(* IEC 61131-3 sources: PLC_ST_Simulator/, 2 files *)

(* ---- Saege_CODESYS.st ---- *)
VAR_GLOBAL
    E0  : BOOL;  (* S0  Rohr an Anschlag 1 *)
    E1  : BOOL;  (* S1  Rohr an Anschlag 2 *)
    E2  : BOOL;  (* S2  gespannt *)
    E3  : BOOL;  (* S3  entspannt *)
    E4  : BOOL;  (* S4  Säge oben *)
    E5  : BOOL;  (* S5  Säge unten *)
    E6  : BOOL;  (* S6  Anschlag 1 oben *)
    E7  : BOOL;  (* S7  Anschlag 1 unten *)
    E8  : BOOL;  (* S8  EIN *)
    E9  : BOOL;  (* S9  AUS, Öffner *)
    E10 : BOOL;  (* S10 Start *)
    E11 : BOOL;  (* S11 Stopp, Öffner *)
    E12 : BOOL;  (* S12 Anschlag 2 oben *)
    E13 : BOOL;  (* S13 Anschlag 2 unten *)
    E14 : BOOL;  (* S14 dickes Rohr *)
    E15 : BOOL;  (* S15 dünnes Rohr *)
    WST_ABTRANSPORT      : BOOL;  (* B1 *)
    mot_schutz_saege     : BOOL;  (* F1..F5 Öffner *)
    mot_schutz_rolle1    : BOOL;
    mot_schutz_rolle2    : BOOL;
    mot_schutz_anschlag1 : BOOL;
    mot_schutz_anschlag2 : BOOL;

    SAEGE_RUNTER     : BOOL;  (* A1 *)
    SAEGE_HOCH       : BOOL;  (* A2 *)
    SPANNEN          : BOOL;  (* A3 *)
    ENTSPANNEN       : BOOL;  (* A4 *)
    SAEGE_ANTRIEB    : BOOL;  (* K1 *)
    ROLLE_1          : BOOL;  (* K2 *)
    ROLLE_2          : BOOL;  (* K3 *)
    ANSCHLAG1_HOCH   : BOOL;  (* K4 *)
    ANSCHLAG1_RUNTER : BOOL;  (* K5 *)
    ANSCHLAG2_HOCH   : BOOL;  (* K6 *)
    ANSCHLAG2_RUNTER : BOOL;  (* K7 *)
END_VAR

FUNCTION_BLOCK FB_Betriebsart
VAR_OUTPUT
    xEin      : BOOL;
    xAuto     : BOOL;
    xStoerung : BOOL;
END_VAR

xStoerung := NOT (mot_schutz_saege AND mot_schutz_rolle1 AND mot_schutz_rolle2
                  AND mot_schutz_anschlag1 AND mot_schutz_anschlag2);

IF E8 THEN xEin := TRUE;END_IF
IF NOT E9 OR xStoerung THEN xEin := FALSE; END_IF

(* Stopp: laufendes Rohr wird fertig bearbeitet *)
IF E10 AND xEin THEN xAuto := TRUE; END_IF
IF NOT E11 OR NOT xEin THEN xAuto := FALSE; END_IF
END_FUNCTION_BLOCK

PROGRAM SFC_Saege
VAR_INPUT
    xAuto      : BOOL;
    xB1_Flanke : BOOL;
    xReset     : BOOL;   (* zurueck in Grundstellung S1 *)
END_VAR
VAR
    iStep     : INT := 1;
    iStepOld  : INT := 0;
    xNeu      : BOOL;    (* Schritt wurde in diesem Zyklus betreten *)
    xDuenn    : BOOL;
    xDick     : BOOL;
    iSoll     : INT;
    iZaehler  : INT;
    xK1, xK2, xK3, xK5, xK7 : BOOL;
    xAbtransport : BOOL;
    xA1, xA2, xA3, xA4 : BOOL;
END_VAR

(* Reset *)
IF xReset THEN
    iStep    := 1;
    iZaehler := 0;
    xDuenn   := FALSE;
    xDick    := FALSE;
END_IF

xNeu     := (iStep <> iStepOld);
iStepOld := iStep;
(* Start *)
IF xNeu THEN
    CASE iStep OF
        2:  (* ACT_Rohrtyp *)
            xDuenn := E15;
            xDick  := E14 AND NOT E15;
            IF xDuenn THEN iSoll := 4; ELSE iSoll := 3; END_IF
        10: (* ACT_Zaehlen *)
            iZaehler := iZaehler + 1;
        11: (* ACT_Ruecksetzen *)
            iZaehler := 0;
            xDuenn   := FALSE;
            xDick    := FALSE;
    END_CASE
END_IF

(*Schrittekette *)
CASE iStep OF
    1:  IF xAuto AND E3 AND E4 AND E6 AND E12 AND (E14 OR E15) THEN iStep := 2;  END_IF
    2:  IF xDuenn THEN iStep := 3;
        ELSIF xDick THEN iStep := 4; END_IF
    3:  IF E7  THEN iStep := 5; END_IF
    4:  IF E13 THEN iStep := 5; END_IF
    5:  IF (xDuenn AND E0) OR (xDick AND E1) THEN iStep := 6; END_IF
    6:  IF E2  THEN iStep := 7; END_IF
    7:  IF E5  THEN iStep := 8; END_IF
    8:  IF E4  THEN iStep := 9; END_IF
    9:  IF E3  THEN iStep := 10; END_IF
    10: IF WST_ABTRANSPORT AND E6 AND E12 THEN
            IF iZaehler < iSoll THEN
                IF xDuenn THEN iStep := 3; ELSE iStep := 4; END_IF
            ELSE
                iStep := 11;
            END_IF
        END_IF
    11: IF xB1_Flanke THEN iStep := 1; END_IF
END_CASE

(* Schrittverriegelungen*)
xK1          := (iStep = 7) OR (iStep = 8);
xK2          := (iStep = 5) OR (iStep = 11);
xK3          := (iStep = 5) OR (iStep = 10) OR (iStep = 11);
xK5          := (iStep = 3);
xK7          := (iStep = 4);
xA1          := (iStep = 7);
xA2          := (iStep = 8);
xA3          := (iStep = 6);
xA4          := (iStep = 9);
xAbtransport := (iStep = 10);
END_PROGRAM

PROGRAM PRG_Ausgaenge
VAR_INPUT
    xFreigabe : BOOL;
END_VAR

ROLLE_1          := xFreigabe AND SFC_Saege.xK2 AND E3;
ROLLE_2          := xFreigabe AND SFC_Saege.xK3;
SPANNEN          := xFreigabe AND SFC_Saege.xA3 AND NOT SFC_Saege.xA4;
ENTSPANNEN       := xFreigabe AND SFC_Saege.xA4 AND E4;
SAEGE_ANTRIEB    := xFreigabe AND SFC_Saege.xK1 AND E2;
SAEGE_RUNTER     := xFreigabe AND SFC_Saege.xA1 AND E2 AND NOT SFC_Saege.xA2;
SAEGE_HOCH       := xFreigabe AND SFC_Saege.xA2;
ANSCHLAG1_HOCH   := xFreigabe AND SFC_Saege.xAbtransport AND SFC_Saege.xDuenn;
ANSCHLAG2_HOCH   := xFreigabe AND SFC_Saege.xAbtransport AND SFC_Saege.xDick;
ANSCHLAG1_RUNTER := xFreigabe AND SFC_Saege.xK5 AND NOT ANSCHLAG1_HOCH;
ANSCHLAG2_RUNTER := xFreigabe AND SFC_Saege.xK7 AND NOT ANSCHLAG2_HOCH;
END_PROGRAM

PROGRAM PLC_PRG
VAR
    fbBetriebsart : FB_Betriebsart;
    rtB1          : R_TRIG;
END_VAR

fbBetriebsart();
rtB1(CLK := WST_ABTRANSPORT);

SFC_Saege(xAuto := fbBetriebsart.xAuto, xB1_Flanke := rtB1.Q, xReset := NOT fbBetriebsart.xEin);

PRG_Ausgaenge(xFreigabe := fbBetriebsart.xEin AND NOT fbBetriebsart.xStoerung);
END_PROGRAM

(* ---- Saege_Anlage.st ---- *)
(* ============================================================
   Anlagenmodell Rohrsäge  –  läuft im Simulator in jedem Zyklus
   VOR dem SPS-Programm und bildet die Sensoren (E0..E15, B1)
   aus den Ausgängen (A1..A4, K1..K7) nach.

   Geometrie (mm, ab Sägeblatt):  Anschlag 1 = 300, Anschlag 2 = 500,
   Lichtschranke B1 = 1500.  Rohrlänge 1700 mm.
   ============================================================ *)

PROGRAM SIM_Saege
VAR_INPUT
    xNaechstesDick : BOOL := FALSE;   (* Typ des nächsten Rohres *)
    xNachladen     : BOOL := TRUE;    (* automatisch neues Rohr auflegen *)
END_VAR
VAR_OUTPUT
    iSchnitte      : INT;             (* Anzahl Schnitte gesamt *)
    iAbtransport   : INT;             (* Teile, die die Anlage verlassen haben *)
    iRohre         : INT;             (* aufgelegte Rohre *)
    xKollision     : BOOL;            (* mechanische Kollision erkannt *)
    sKollision     : STRING;
END_VAR
VAR CONSTANT
    POS_A1   : REAL := 300.0;
    POS_A2   : REAL := 500.0;
    POS_B1   : REAL := 1500.0;
    ROHR_LEN : REAL := 1700.0;
    V_ROLLE  : REAL := 0.5;     (* mm/ms *)
    V_SAEGE  : REAL := 0.1;     (* %/ms  -> 1 s Hub *)
    V_SPANN  : REAL := 0.4;     (* %/ms  -> 250 ms *)
    V_ANSCHL : REAL := 0.25;    (* %/ms  -> 400 ms *)
    MAX_TEILE : INT := 8;
END_VAR
VAR
    xInit      : BOOL;
    tLast      : TIME;
    dt         : REAL;
    rSaege     : REAL := 100.0;  (* 100 = oben, 0 = unten *)
    rSpann     : REAL := 0.0;    (* 0 = entspannt, 100 = gespannt *)
    rAnschlag1 : REAL := 0.0;    (* 0 = oben, 100 = unten *)
    rAnschlag2 : REAL := 0.0;
    xRohrDick  : BOOL;
    rRohrFront : REAL;           (* Rohranfang hinter dem Sägeblatt *)
    rRohrLen   : REAL;           (* Restlänge auf der Zuführung *)
    aFront     : ARRAY[1..8] OF REAL;   (* abgesägte Teile auf Rollenbahn 2 *)
    aLen       : ARRAY[1..8] OF REAL;
    nTeile     : INT;
    xGeschnitten : BOOL;
    tonLaden   : TON;
    i, k       : INT;
    rWeg, rHinten : REAL;
END_VAR

(* ---------- Initialisierung beim ersten Zyklus ---------- *)
IF NOT xInit THEN
    xInit := TRUE;
    tLast := TIME();
    E9 := TRUE;  E11 := TRUE;   (* Öffner nicht betätigt *)
    mot_schutz_saege := TRUE;  mot_schutz_rolle1 := TRUE;  mot_schutz_rolle2 := TRUE;
    mot_schutz_anschlag1 := TRUE;  mot_schutz_anschlag2 := TRUE;
END_IF
dt := TIME_TO_REAL(TIME() - tLast);
tLast := TIME();

(* ---------- Säge ---------- *)
IF SAEGE_RUNTER AND NOT SAEGE_HOCH THEN
    rSaege := MAX(0.0, rSaege - V_SAEGE * dt);
ELSIF SAEGE_HOCH AND NOT SAEGE_RUNTER THEN
    rSaege := MIN(100.0, rSaege + V_SAEGE * dt);
END_IF
IF rSaege < 60.0 AND rRohrLen > 0.0 AND NOT SAEGE_ANTRIEB AND NOT xKollision THEN
    xKollision := TRUE;  sKollision := 'Säge fährt ohne Antrieb ins Rohr';
END_IF
IF rSaege < 60.0 AND rRohrLen > 0.0 AND rSpann < 100.0 AND NOT xKollision THEN
    xKollision := TRUE;  sKollision := 'Sägen ohne gespanntes Rohr';
END_IF

(* ---------- Spannbacken ---------- *)
IF SPANNEN AND NOT ENTSPANNEN THEN
    rSpann := MIN(100.0, rSpann + V_SPANN * dt);
ELSIF ENTSPANNEN AND NOT SPANNEN THEN
    rSpann := MAX(0.0, rSpann - V_SPANN * dt);
END_IF

(* ---------- Längenanschläge ---------- *)
IF ANSCHLAG1_RUNTER AND NOT ANSCHLAG1_HOCH THEN rAnschlag1 := MIN(100.0, rAnschlag1 + V_ANSCHL * dt);
ELSIF ANSCHLAG1_HOCH AND NOT ANSCHLAG1_RUNTER THEN rAnschlag1 := MAX(0.0, rAnschlag1 - V_ANSCHL * dt); END_IF
IF ANSCHLAG2_RUNTER AND NOT ANSCHLAG2_HOCH THEN rAnschlag2 := MIN(100.0, rAnschlag2 + V_ANSCHL * dt);
ELSIF ANSCHLAG2_HOCH AND NOT ANSCHLAG2_RUNTER THEN rAnschlag2 := MAX(0.0, rAnschlag2 - V_ANSCHL * dt); END_IF

(* Anschlag fährt auf ein Teil, das unter ihm liegt? *)
FOR i := 1 TO nTeile DO
    rHinten := aFront[i] - aLen[i];
    IF ANSCHLAG1_RUNTER AND rHinten < POS_A1 - 1.0 AND aFront[i] > POS_A1 + 1.0 AND NOT xKollision THEN
        xKollision := TRUE;  sKollision := 'Anschlag 1 fährt auf ein Teil';
    END_IF
    IF ANSCHLAG2_RUNTER AND rHinten < POS_A2 - 1.0 AND aFront[i] > POS_A2 + 1.0 AND NOT xKollision THEN
        xKollision := TRUE;  sKollision := 'Anschlag 2 fährt auf ein Teil';
    END_IF
END_FOR

IF ANSCHLAG1_RUNTER AND rRohrLen > 0.0 AND rRohrFront > POS_A1 + 1.0 AND NOT xKollision THEN
    xKollision := TRUE;  sKollision := 'Anschlag 1 fährt auf das Rohr';
END_IF
IF ANSCHLAG2_RUNTER AND rRohrLen > 0.0 AND rRohrFront > POS_A2 + 1.0 AND NOT xKollision THEN
    xKollision := TRUE;  sKollision := 'Anschlag 2 fährt auf das Rohr';
END_IF

(* ---------- Rohr auf der Zuführung (Rollenbahn 1) ---------- *)
IF ROLLE_1 AND rRohrLen > 0.0 THEN
    IF rSpann > 0.0 THEN
        IF NOT xKollision THEN xKollision := TRUE; sKollision := 'Vorschub gegen gespanntes Rohr'; END_IF
    ELSE
        rWeg := V_ROLLE * dt;
        rRohrFront := rRohrFront + rWeg;
        IF rAnschlag1 > 0.0 AND rRohrFront - rWeg <= POS_A1 + 0.01 THEN rRohrFront := MIN(rRohrFront, POS_A1); END_IF
        IF rAnschlag2 > 0.0 AND rRohrFront - rWeg <= POS_A2 + 0.01 THEN rRohrFront := MIN(rRohrFront, POS_A2); END_IF
        (* Rohrende hat die Säge passiert -> Reststück auf Rollenbahn 2 *)
        IF rRohrFront >= rRohrLen AND nTeile < MAX_TEILE THEN
            nTeile := nTeile + 1;
            aFront[nTeile] := rRohrFront;  aLen[nTeile] := rRohrLen;
            rRohrLen := 0.0;  rRohrFront := 0.0;
        END_IF
    END_IF
END_IF

(* ---------- Schnitt ---------- *)
IF SAEGE_ANTRIEB AND rSaege <= 0.0 AND rSpann >= 100.0 AND NOT xGeschnitten AND rRohrFront > 0.0 AND nTeile < MAX_TEILE THEN
    xGeschnitten := TRUE;
    iSchnitte := iSchnitte + 1;
    nTeile := nTeile + 1;
    aFront[nTeile] := rRohrFront;  aLen[nTeile] := rRohrFront;
    rRohrLen := rRohrLen - rRohrFront;
    rRohrFront := 0.0;
END_IF
IF rSaege >= 100.0 THEN xGeschnitten := FALSE; END_IF

(* ---------- Teile auf Rollenbahn 2 ---------- *)
IF ROLLE_2 THEN
    rWeg := V_ROLLE * dt;
    FOR i := 1 TO nTeile DO
        aFront[i] := aFront[i] + rWeg;
        IF rAnschlag1 > 0.0 AND aFront[i] - rWeg <= POS_A1 + 0.01 THEN aFront[i] := MIN(aFront[i], POS_A1); END_IF
        IF rAnschlag2 > 0.0 AND aFront[i] - rWeg <= POS_A2 + 0.01 THEN aFront[i] := MIN(aFront[i], POS_A2); END_IF
    END_FOR
END_IF
(* Teile, die die Rollenbahn verlassen haben, entfernen *)
i := 1;
WHILE i <= nTeile DO
    IF aFront[i] - aLen[i] > POS_B1 + 300.0 THEN
        FOR k := i TO nTeile - 1 DO
            aFront[k] := aFront[k + 1];  aLen[k] := aLen[k + 1];
        END_FOR
        nTeile := nTeile - 1;
        iAbtransport := iAbtransport + 1;
    ELSE
        i := i + 1;
    END_IF
END_WHILE

(* ---------- Rohr nachladen ---------- *)
tonLaden(IN := xNachladen AND rRohrLen <= 0.0 AND NOT ROLLE_1, PT := T#1s);   (* Werker legt nur bei stehender Bahn auf *)
IF tonLaden.Q THEN
    rRohrLen := ROHR_LEN;  rRohrFront := 0.0;
    xRohrDick := xNaechstesDick;
    iRohre := iRohre + 1;
END_IF

(* ---------- Sensoren ---------- *)
E0  := rRohrLen > 0.0 AND rAnschlag1 >= 100.0 AND rRohrFront >= POS_A1 - 0.5;
E1  := rRohrLen > 0.0 AND rAnschlag2 >= 100.0 AND rRohrFront >= POS_A2 - 0.5;
E2  := rSpann >= 100.0;
E3  := rSpann <= 0.0;
E4  := rSaege >= 100.0;
E5  := rSaege <= 0.0;
E6  := rAnschlag1 <= 0.0;
E7  := rAnschlag1 >= 100.0;
E12 := rAnschlag2 <= 0.0;
E13 := rAnschlag2 >= 100.0;
E14 := rRohrLen > 0.0 AND xRohrDick;
E15 := rRohrLen > 0.0 AND NOT xRohrDick;
WST_ABTRANSPORT := FALSE;
FOR i := 1 TO nTeile DO
    IF aFront[i] >= POS_B1 AND aFront[i] - aLen[i] <= POS_B1 THEN WST_ABTRANSPORT := TRUE; END_IF
END_FOR
END_PROGRAM
